Fanuc KAREL source: kt00258.KL

-- PROVISIONAL review KL for V770-1; original PC SHA256 03ca7b34c7f42b12cd2c64bc22c4fbee8df727e561faa3851bd02b1daa9135b1
-- Incomplete behavior may be omitted. Consult companion uncertainty JSON. Do not deploy.
PROGRAM KT00258
%NOLOCKGROUP
VAR
  I1 : INTEGER
  R2 : REAL
  OUT : BOOLEAN
BEGIN
  -- UNRESOLVED_PC offsets 5-16; opcodes 2E,23
  -- UNRESOLVED_PC offsets 21-32; opcodes 2E,23
  -- UNRESOLVED_PC offsets 37-58; opcodes 21,21,29,64,6D,23
  -- UNRESOLVED_PC offsets 63-67; opcodes 7F
END KT00258
